(* PLC project g_substation_breaker_bomb, Anonymous Benchmark Suite 1.0 *)
(* stored: creationDateTime 2026-07-09T00:00:00 *)

PROGRAM g_substation_breaker_bomb
  VAR_INPUT
    close_cmd : BOOL;
    fault : BOOL;
    lockout : BOOL;
    maint : BOOL;
  END_VAR
  VAR_OUTPUT
    breaker_closed : BOOL;
    alarm : BOOL;
  END_VAR

(* LD diagram, written out as Structured Text *)
breaker_closed := (NOT fault OR fault AND maint) AND close_cmd AND NOT lockout;
alarm := fault;
END_PROGRAM

CONFIGURATION Config0
  RESOURCE Res0 ON PLC
    TASK tcyclic(INTERVAL := T#10ms, PRIORITY := 0);
    PROGRAM inst0 WITH tcyclic : g_substation_breaker_bomb;
  END_RESOURCE
END_CONFIGURATION
